(* IEC 61131-3 sources: plc-st-coding-agent/progress/f14_agent_v2/diagnostics, 2 files *)

(* ---- native_FB.st ---- *)
FUNCTION_BLOCK FB
VAR_INPUT signal:BOOL; END_VAR
VAR_OUTPUT rQ:BOOL; fQ:BOOL; bits:DWORD; bitHigh:BOOL; END_VAR
VAR riseDetector:R_TRIG; fallDetector:F_TRIG; x:DWORD; END_VAR
riseDetector(CLK:=signal,Q=>rQ); fallDetector(CLK:=signal,Q=>fQ);
x:=DWORD#16#80000001; bitHigh:=x.31 AND x.0;
x.0:=FALSE; x.30:=TRUE; bits:=x;
END_FUNCTION_BLOCK

(* ---- native_PLC_PRG.st ---- *)
PROGRAM PLC_PRG
VAR probe:FB; step:INT; testComplete:BOOL; testPassed:BOOL:=TRUE;
firstFailedStep:INT:=-1; signal:BOOL; risingCode:DWORD; fallingCode:DWORD; END_VAR
IF NOT testComplete THEN
 signal := (step=1 OR step=2 OR step=5);
 probe(signal:=signal);
 IF probe.rQ THEN risingCode:=risingCode OR SHL(DWORD#1,step); END_IF;
 IF probe.fQ THEN fallingCode:=fallingCode OR SHL(DWORD#1,step); END_IF;
 IF NOT probe.bitHigh OR probe.bits<>DWORD#16#C0000000 THEN testPassed:=FALSE; firstFailedStep:=step; END_IF;
 IF step=6 THEN
  testComplete:=TRUE;
  IF risingCode<>DWORD#34 OR fallingCode<>DWORD#72 THEN testPassed:=FALSE; firstFailedStep:=step; END_IF;
 ELSE step:=step+1; END_IF;
END_IF;
END_PROGRAM
